(* IEC 61131-3 sources: lasal-git-demo/CPU/LasalDemoProject/Class/ECAT_Master_Base (part 2) *)

#ifdef ECAT_DEBUG_TIMEMEASURE2
          pCTI^.ud_TimePre := OS_GETMICROSEC() - udTimeMarkus;
          if pCTI^.ud_TimePre < pCTI^.ud_TimePreMin then
            pCTI^.ud_TimePreMin := pCTI^.ud_TimePre;
          end_if;
          if pCTI^.ud_TimePre > pCTI^.ud_TimePreMax then
            pCTI^.ud_TimePreMax := pCTI^.ud_TimePre;
          end_if;
#endif
        else

          //Check the process state if we need to raise an error
          dTriggerFrameError := ProcessFrameErrorCheck(pCTI^.ecatm_cycctx^.prcstatus);

          //Check if we need to trigger an error
          if dTriggerFrameError then
            ClassState := _WrongRunStatus;

            bd_LogRtMessagesInCy.PostIt.CycPrcStatus  := TRUE;
            bd_LogRtMessagesInCy.aLogValue1[14]       := pCTI^.ecatm_cycctx^.prcstatus;

            if bd_Flags.bIsRequired then
              CrashThisTime := TRUE;
              sigclib_sprintfST(pd:=#aCrashMessage[0], format:="Ethercat: Error (Invalid frame) Status 0x%X", p0:=#pCTI^.ecatm_cycctx^.prcstatus);
            end_if;
          end_if;
        end_if;

        MissedFrameCounter := sDebugCounters.udConsecutiveMissingFrameCounter;

      end_if;

    else

      sDebugCounters.udInvalidcycctx += 1;

      //Cyclic Context is not valid until EtherCAT State is OP or higher
      if EtherCATState >= ECAT_STATE_OP then
        //Cyclic context is invalid although the EtherCAT State is higher or equal than SAFEOP --> SET Error
        ClassState    := _WrongRunStatus;

        bd_LogRtMessagesInCy.PostIt.InvalidCycctx := TRUE;

        if bd_Flags.bIsRequired then
          CrashThisTime := TRUE;
          _strcpy(dest:=#aCrashMessage[0], src:="EtherCAT: Invalid Cycctx");
        end_if;
      end_if;

    end_if;

  else

    if retcode < ECATM_OK then  // retcode may be of type t_e_st_ecatm_evtc in this case we need unlock
      bNoUnlock := TRUE;
    end_if;

    sDebugCounters.udInvalidRetCodeUpdateCycPre += 1;

    CrashThisTime := UpdateCycRetcodeHandling(retcode:=retcode, pCrashMessage:=#aCrashMessage[0]);

  end_if;

  // Always Call to unlock cycctx
  if ( (pCTI^.bPostScanActive) = FALSE |    // Postscan call needed to unlock ecatm_cycctx
       (EtherCATState < ECAT_STATE_OP) |    // If EtherCATState = OP then unlock is done in postscan
       ((ClassState <> _ClassOk) & (bNoUnlock = FALSE)) ) then     // Unlock on Error, Postscan is no longer called in this state

#ifdef ECAT_TRACE_VIEW_LOG
    OS_MakeTraceEntry(pSystrace, HWCONTROL_SYSTRACE_TYPE, ECAT_SYSTRACE_PRESCAN_UPDATECYC_UNLOCK,pCTI^.udCycTaskId);
#endif

    retcode := OS_ECATM_UpdateCyc(pECAT, ecatmhdl, pCTI^.udCycTaskId, LSL_ECATM_POST_CYC_TASK, #pCTI^.ecatm_cycctx,0);
    if retcode <> ECATM_OK then

      //Invalid retcode, raise error
      sDebugCounters.udInvalidRetCodeUpdateCycPost += 1;

      CrashThisTime := UpdateCycRetcodeHandling(retcode:=retcode, pCrashMessage:=#aCrashMessage[0]);

    end_if;
  end_if;

  if CrashThisTime then
    // if a required module is not available or doesn't work properly, the system should crash
    OS_ECATM_raise_error(pECAT,0,#aCrashMessage[0]);
  end_if;

END_FUNCTION

FUNCTION VIRTUAL GLOBAL ECAT_Master_Base::UpdateRtPostScan
  VAR_INPUT
    pCTI 	: ^t_s_CycTaskInfo;
  END_VAR
  VAR
    i               : UDINT;
    pCallbackData   : ^t_s_MapPDOData;
    CrashThisTime   : BOOL;
    aCrashMessage   : ARRAY [0..255] OF CHAR;
    retcode         : DINT;
    dTriggerFrameError  : DINT;
    prcstatus       : UDINT;
#ifdef ECAT_DEBUG_TIMEMEASURE2
    udTimeMarkus : UDINT;
#endif
  END_VAR

  CrashThisTime   := FALSE; // init with false

  //Check if we have postscan callbacks and a valid frame
  if pCTI^.noPostCallbacks & pCTI^.ecatm_cycctx then

    pCallbackData := pCTI^.pPostCallbacks;
    prcstatus := pCTI^.ecatm_cycctx^.prcstatus; // Save prcstatus as it is checked more than once
    if (prcstatus AND ECATM_PRCSTAT_ST_FRAME_NOT_SENT) = 0 then // ECATM_PRCSTAT_ST_FRAME_NOT_SENT: The link layer driver failed to send the last TX frame.
                                                                //                                  The frame is still owned by the hardware of the MAC.
                                                                //                                  THE APPLICATION SHALL NOT ALTER THE TRANSMIT FRAME!
                                                                // Check the sample-simple and sample-all implementation for usaage and compatibility patch.
                                                                // See ECATM_Programmers_Guide and ECATM_Reference_Manual for detailed information

#ifdef ECAT_DEBUG_TIMEMEASURE2
      udTimeMarkus := OS_GETMICROSEC();
#endif

      //Go through all installed callbacks from the slave modules HWK to fetch the data and copy it to the transmit frame.
      for i := 1 to pCTI^.noPostCallbacks do

        if pCallbackData^.pEtherCatState^ >= ECAT_STATE_OP then

#ifdef ECAT_TRACE_VIEW_LOG
            OS_MakeTraceEntry(pSystrace, HWCONTROL_SYSTRACE_TYPE, ECAT_SYSTRACE_POSTSCAN_CALLBACKS,pCTI^.udCycTaskId OR (i SHL 16));
#endif

          pCallbackData^.pCallBack$ECAT_MapPDOData(pCallbackData^.pThis, pCTI^.ecatm_cycctx, pCallbackData^.noData, pCallbackData^.iovar, pCallbackData^.pData);
        end_if;

        pCallbackData += sizeof(t_s_MapPDOData);
      end_for;

#ifdef ECAT_DEBUG_TIMEMEASURE2
      pCTI^.ud_TimePost := OS_GETMICROSEC() - udTimeMarkus;
      if pCTI^.ud_TimePost < pCTI^.ud_TimePostMin then
        pCTI^.ud_TimePostMin := pCTI^.ud_TimePost;
      end_if;
      if pCTI^.ud_TimePost > pCTI^.ud_TimePostMax then
        pCTI^.ud_TimePostMax := pCTI^.ud_TimePost;
      end_if;
#endif
    end_if;

    if (prcstatus AND ECATM_PRCSTAT_ST_MASK_ERROR_OR_WARN) then

      //Check only if no Prescan is used - otherwise this check is done in prescan
      if pCTI^.noPreCallbacks = 0 then

        //Check the process state if we need to raise an error
        dTriggerFrameError := ProcessFrameErrorCheck(prcstatus);

        if dTriggerFrameError then
          ClassState := _WrongRunStatus;

          bd_LogRtMessagesInCy.PostIt.CycPrcStatus  := TRUE;
          bd_LogRtMessagesInCy.aLogValue1[14]       := prcstatus;

          if bd_Flags.bIsRequired then
            CrashThisTime := TRUE;
            sigclib_sprintfST(pd:=#aCrashMessage[0], format:="Ethercat: Error (Invalid frame) Status 0x%X", p0:=#prcstatus);
          end_if;
        end_if;
      end_if;
    end_if;

    MissedFrameCounter := sDebugCounters.udConsecutiveMissingFrameCounter;

  end_if;

#ifdef ECAT_TRACE_VIEW_LOG
  OS_MakeTraceEntry(pSystrace, HWCONTROL_SYSTRACE_TYPE, ECAT_SYSTRACE_POSTSCAN_UPDATECYC,pCTI^.udCycTaskId);
#endif

  // Always Call to unlock cyctx
  retcode := OS_ECATM_UpdateCyc(pECAT, ecatmhdl, pCTI^.udCycTaskId, LSL_ECATM_POST_CYC_TASK, #pCTI^.ecatm_cycctx,0);

  if udDisconnectEventTime then
    udDisconnectEventTime := 0;
    ClassState := _NoHardware;
    EtherCATState := ECAT_STATE_INIT;
    NewMasterEtherCATState  := ECAT_STATE_INIT;
    InitSSW := _Wait4EcatLink;
  end_if;

  if retcode <> ECATM_OK then
    //Invalid retcode, raise error
    sDebugCounters.udInvalidRetCodeUpdateCycPost += 1;

    CrashThisTime := UpdateCycRetcodeHandling(retcode:=retcode, pCrashMessage:=#aCrashMessage[0]);

  end_if;

  if CrashThisTime then
    // if a required module is not available or doesn't work properly, the system should crash
    OS_ECATM_raise_error(pECAT,0,#aCrashMessage[0]);
  end_if;

END_FUNCTION

FUNCTION VIRTUAL ECAT_Master_Base::UpdateCycRetcodeHandling
  VAR_INPUT
    retcode 	: DINT;
    pCrashMessage : ^Char;
  END_VAR
  VAR_OUTPUT
    bFatalError : BOOL;
  END_VAR

  bFatalError := FALSE;

  //Difference the single errors
  case retcode of
    //*****************************************************************************
    ECATM_TIMING_ERROR_1:

      //No Data available at send time (last cycle)
      ClassState := _TimesliceErrorIRQ;
      bd_LogRtMessagesInCy.PostIt.TimingError_1 := TRUE;

      if bd_Flags.bIsRequired then
        bFatalError := TRUE;
        _strcpy(dest:=pCrashMessage, src:="No Data available at Send time (TimeSliceErrorIRQ)");
      end_if;

    //*****************************************************************************
    ECATM_TIMING_ERROR_2:

      //Time since tick is at call of UpdateCyc(Pre) higher than allowed from the IsoStartPoint
      ClassState := _TimesliceErrorIRQ;
      bd_LogRtMessagesInCy.PostIt.TimingError_2 := TRUE;

      if bd_Flags.bIsRequired then
        bFatalError := TRUE;
        _strcpy(dest:=pCrashMessage, src:="Time since tick is at call of UpdateCyc(Pre) higher than allowed from the IsoStartPoint (TimeSliceErrorIRQ)");
      end_if;

    //*****************************************************************************
    ECATM_DATA_NOT_SENT:

      //Data was not sent at the time UpdateCyc was called with (Pre)
      ClassState := _TimesliceError;
      bd_LogRtMessagesInCy.PostIt.DataNotSent := TRUE;

      if bd_Flags.bIsRequired then
        bFatalError := TRUE;
        _strcpy(dest:=pCrashMessage, src:="Data was not sent at the time UpdateCyc was called with (Pre) (TimeSliceError)");
      end_if;

    //*****************************************************************************
    else

      if retcode = ECATM_EVTC_MST_DEACTIVATED$DINT & InitSSW <> _InitFinished then
        //Ignore master deactivated error during initialisation (maybe master is not activated yet (takes a while in OS)

      else
        ClassState := _ManagerError;
        bd_LogRtMessagesInCy.PostIt.UnknownError := TRUE;
        bd_LogRtMessagesInCy.aLogValue1[4] := (ABS(retcode))$UDINT;
        if bd_Flags.bIsRequired then
          bFatalError := TRUE;
          sigclib_sprintfST(pd:=pCrashMessage, format:="Unknown Error in EtherCAT handling occured: %d", p0:=#retcode);
        end_if;
      end_if;

    //*****************************************************************************
  end_case;

END_FUNCTION

FUNCTION VIRTUAL GLOBAL ECAT_Master_Base::SoftwareVersion::Read
  VAR_OUTPUT
    output (EAX) 	: UDINT;
  END_VAR

  SoftwareVersion := strSoftwareVersion.Data.Read();
  output := SoftwareVersion;

END_FUNCTION

FUNCTION VIRTUAL GLOBAL ECAT_Master_Base::SoftwareVersion::Write
  VAR_INPUT
    input (EAX) 	: UDINT;
  END_VAR
  VAR_OUTPUT
    result (EAX) 	: UDINT;
  END_VAR

  SoftwareVersion := input;
  result := (strSoftwareVersion.Data.Write(SoftwareVersion))$UDINT;

END_FUNCTION

FUNCTION VIRTUAL GLOBAL ECAT_Master_Base::CyWork
  VAR_INPUT
    EAX 	: UDINT;
  END_VAR
  VAR_OUTPUT
    state (EAX) 	: UDINT;
  END_VAR
  VAR
    pCurrentSlave : ^t_sSlaveInfo;
    i             : UDINT;
    _Para         : CmdStruct;
    _Result       : Results;
    RetCodeIPR    : iprStates;
    b_ModulInitComplete   : BOOL;
    TmpRequest    : BDINT;
    retCode       : DINT;
  END_VAR

  case InitSSW of
//**********************************************************************************************************************************************************
    t_e_InitSSW::_StartInit:

#ifdef ECAT_TRACE_VIEW_LOG
      OS_MakeTraceEntry(pSystrace, HWCONTROL_SYSTRACE_TYPE, ECAT_SYSTRACE_POSTINIT_START_INIT,0);
#endif

      // remember when we started (for timeout and init time measure)
      udInitStartTime := ops.tAbsolute;

      // check if we had an error before
      if InitError <> _ClassOk then
        // we already have a log entry from the init
        ClassState := InitError;
        ErrorInitStep := InitSSW;
        InitSSW := _PrepareError;
        EtherCATState := ECAT_STATE_NONE;
        return;
      end_if;

      // Check if post init needs to be extended
      if StateTransitionTimeout.Read() > POST_INIT_TIMEOUT then

        ExtendPostInitTime(AdditionalTime:=StateTransitionTimeout);

      end_if;

      InitSSW := _Wait4ECATLink;

//**********************************************************************************************************************************************************
    t_e_InitSSW::_Wait4ECATLink:

      retCode := OS_ECATM_NET_GET_STATUS(pECAT, ecatmhdl, #snetStatus);

      if retCode then
        LogValue("@0563 (ECAT_Master_Base::CyWork) Failed to get ECAT Link Status. Return Code: 0x{0} via InitModule-Interface", retCode$UDINT);

        ErrorInitStep := InitSSW;
        InitSSW := _PrepareError;
        ClassState := InitError    := _ManagerError;
        EtherCATState := ECAT_STATE_NONE;

        return;
      end_if;

      if snetStatus.flags.ECATM_NET_STATUS_MST_LINK_DOWN = FALSE then

#ifdef ECAT_DEBUG_EVENT_CALLBACKS
        LogValue("ECAT-DEBUG: Link found after 0x{0}ms", (ops.tAbsolute-udInitStartTime));
#endif

        //ClassState is set to NoHardware at DisconnectEvent -> Set back to _ClassOk to ensure that the Realtime functions are called
        ClassState := _ClassOk;

        //Go on and call the connect event methods
        InitSSW := _CallConnectEventOfModules;
      elsif ( (bd_Flags.bDisableWait4LinkTimeOut = FALSE) &
              (ops.tAbsolute - udInitStartTime) > GetWait4LinkTimeout()) then

        ErrorInitStep := InitSSW;
        InitSSW       := _PrepareError;
        ClassState    := InitError     := _ManagerError;
        EtherCATState := ECAT_STATE_NONE;
        LogError("@067B (ECAT_Master_Base::CyWork) Master Link Down (Timeout)! Unable to continue with Initialisation.");

      end_if;

//**********************************************************************************************************************************************************
    t_e_InitSSW::_CallConnectEventOfModules:

      //Call the Connect Event of every slave
      if sSlaveInfo.udMaxSlaves then
        pCurrentSlave := sSlaveInfo.pSlaves; //Point to current slave
        for i:=0 to sSlaveInfo.udMaxSlaves-1 do
          //Only call module if no error
          if pCurrentSlave^.pThis & pCurrentSlave^.pThis^.EtherCATState <> ECAT_STATE_NONE then
            pCurrentSlave^.pThis^.ConnectEvent();
          end_if;
          pCurrentSlave += sizeof(t_sSlaveInfo);
        end_for;
      end_if;

      InitSSW := _PrepareNextEtherCATState;

//**********************************************************************************************************************************************************
    t_e_InitSSW::_PrepareNextEtherCATState:

      //Go on with next step of initialisation
      InitSSW := _SwitchToNextEtherCATState;
      TmpRequest := 0;

      //Check if any slave needs an InitModule call. Otherwise we can directy request the OP State from the master
      if sSlaveInfo.udMaxSlaves then
        pCurrentSlave := sSlaveInfo.pSlaves; //Point to current slave
        //Call UpdateCy of all logged in slaves
        for i:=0 to sSlaveInfo.udMaxSlaves-1 do
          if pCurrentSlave^.pThis & pCurrentSlave^.bdInitModuleFlags <> ECAT_INIT_MODULE_NO_CALL then
            TmpRequest := TmpRequest OR pCurrentSlave^.bdInitModuleFlags;
          end_if;
          pCurrentSlave += sizeof(t_sSlaveInfo);
        end_for;
      end_if;

      //Determine master state to request (e.g. if no module needs to be called during our InitModulePhase, we can directly request the OP State)
      if (TmpRequest AND ECAT_INIT_MODULE_CALL_INIT) = ECAT_INIT_MODULE_CALL_INIT then
        RequestMasterState := ECAT_STATE_INIT;
      elsif (TmpRequest AND ECAT_INIT_MODULE_CALL_PREOP) = ECAT_INIT_MODULE_CALL_PREOP then
        RequestMasterState := ECAT_STATE_PREOP;
      elsif (TmpRequest AND ECAT_INIT_MODULE_CALL_SAFEOP) = ECAT_INIT_MODULE_CALL_SAFEOP then
        RequestMasterState := ECAT_STATE_SAFEOP;
      else
        //No module needs an InitModule Call
        RequestMasterState := ECAT_STATE_OP;
      end_if;

//**********************************************************************************************************************************************************
    t_e_InitSSW::_SwitchToNextEtherCATState:

      //Set master to determined state
#ifdef ECAT_DEBUG_EVENT_CALLBACKS
      LogValue(pString:="ECAT-DEBUG: Request New ECATMST State: 0x{0}", Value:=RequestMasterState);
#endif
      retcode := OS_ECATM_MST_REQ_STATE(pECAT, ecatmhdl, RequestMasterState, StateTransitionBehaviour);
      if retcode then
        LogValue("@0565 (ECAT_Master_Base::CyWork) Call OS_ECATM_MST_REQ_STATE() Failed with retcode 0x{0}! Unable to continue with Initialisation", ABS(retcode)$UDINT);
        // Disable Class
        ErrorInitStep := InitSSW;
        InitSSW := _PrepareError;
        ClassState := _ManagerError;
        EtherCATState := ECAT_STATE_NONE;
        return;
      end_if;

      udCheckEtherCATStateTime := ops.tAbsolute;
      InitSSW := _CheckEtherCATState;

//**********************************************************************************************************************************************************
    t_e_InitSSW::_CheckEtherCATState:

      //Wait until master is in requested state
      if EtherCATState = RequestMasterState then

#ifdef ECAT_TRACE_VIEW_LOG
        OS_MakeTraceEntry(pSystrace, HWCONTROL_SYSTRACE_TYPE, ECAT_SYSTRACE_POSTINIT_CHECK_ETHERCAT_STATE,EtherCATState$UDINT);
#endif

        //If we are in the requested state go on with InitModule Phase
        InitSSW := _CallInitModule;

        udInitModuleTimeStamp := ops.tAbsolute;
        udInitModuleTimeOut   := GetCallInitModuleTimeout();

      elsif ( (bd_Flags.bDisableStateTransitionTimeout = FALSE) &
              (ops.tAbsolute - udCheckEtherCATStateTime) > StateTransitionTimeout.Read()) then
        LogValue("@0566 (ECAT_Master_Base::CyWork) Timeout while waiting for EtherCATState! EtherCATState: 0x{0}, RequestMasterState: 0x{1}", EtherCATState$UDINT,RequestMasterState$UDINT);
        ErrorInitStep := InitSSW;
        InitSSW := _PrepareError;
        ClassState := _TimeoutInInit;
        EtherCATState := ECAT_STATE_NONE;
        return;
      end_if;

//**********************************************************************************************************************************************************
    t_e_InitSSW::_CallInitModule:

      // preinitialize the complete marker => is resetted if a module has to be initialized
      b_ModulInitComplete := TRUE;

      //Call all slaves (needed for SDO Handling)
      if sSlaveInfo.udMaxSlaves then
        pCurrentSlave := sSlaveInfo.pSlaves; //Point to current slave

        _Para.uiCmd := ECAT_M_CALL_INIT_MODULE;
        _Para.aPara[0]$DINT           := 1;
        _Para.aPara[1]$t_e_ECAT_STATE := EtherCATState;

        //Call UpdateCy of all logged in slaves
        for i:=0 to sSlaveInfo.udMaxSlaves-1 do

          //Check if current module has to be called
          if (pCurrentSlave^.bdInitModuleFlags <> ECAT_INIT_MODULE_NO_CALL) &
            ((pCurrentSlave^.bdInitModuleFinished AND EtherCATState$BDINT) <> EtherCATState$BDINT ) then

            if (EtherCATState = ECAT_STATE_INIT   & ((pCurrentSlave^.bdInitModuleFlags AND ECAT_INIT_MODULE_CALL_INIT)    = ECAT_INIT_MODULE_CALL_INIT))  |
               (EtherCATState = ECAT_STATE_PREOP  & ((pCurrentSlave^.bdInitModuleFlags AND ECAT_INIT_MODULE_CALL_PREOP)   = ECAT_INIT_MODULE_CALL_PREOP)) |
               (EtherCATState = ECAT_STATE_SAFEOP & ((pCurrentSlave^.bdInitModuleFlags AND ECAT_INIT_MODULE_CALL_SAFEOP)  = ECAT_INIT_MODULE_CALL_SAFEOP)) |
               (EtherCATState = ECAT_STATE_OP     & ((pCurrentSlave^.bdInitModuleFlags AND ECAT_INIT_MODULE_CALL_OP)      = ECAT_INIT_MODULE_CALL_OP))
            then
              RetCodeIPR := pCurrentSlave^.pThis^.NewInst(#_Para,#_Result);

#ifdef ECAT_TRACE_VIEW_LOG
              OS_MakeTraceEntry(pSystrace, HWCONTROL_SYSTRACE_TYPE, ECAT_SYSTRACE_POSTINIT_CALL_INITMODULE,i);
#endif
              //Check retcode
              if RetCodeIPR = ERROR then

                LogValue("@0567 (ECAT_Master_Base::CyWork) Failed to initialize EtherCAT Slave 0x{0} via InitModule-Interface", i);

                // Set as finshed so that not required module is not called again and does not spam log
                // Disable Init callbacks for all EtherCAT States
                pCurrentSlave^.bdInitModuleFinished := pCurrentSlave^.bdInitModuleFinished OR ECAT_STATE_INIT$BDINT OR ECAT_STATE_PREOP$BDINT OR ECAT_STATE_SAFEOP$BDINT OR ECAT_STATE_OP$BDINT;

                // if it's an required module => error
                if pCurrentSlave^.bRequired   then
                  SetRequiredError( pTargetThis       := pCurrentSlave^.pThis
                                  , udSlaveIndex      := pCurrentSlave^.udSlaveIndex
                                  , bLogInMethAllowed := TRUE);
                end_if;

              elsif RetCodeIPR = READY then
                pCurrentSlave^.bdInitModuleFinished := pCurrentSlave^.bdInitModuleFinished OR EtherCATState$BDINT;
              else
                b_ModulInitComplete := FALSE; //At least one module is not ready yet --> carry on with ModuleInit phase
              end_if;
            //else
              //Module will be called if the needed EtherCAT State is active
            end_if;
          else
            //Module has no need to be called, just set as finished
            pCurrentSlave^.bdInitModuleFinished := pCurrentSlave^.bdInitModuleFinished OR EtherCATState$BDINT;
          end_if;

          pCurrentSlave += sizeof(t_sSlaveInfo);
        end_for;
      end_if;

      //Check if every module init is finished, go on to next state
      if b_ModulInitComplete = TRUE then

        InitSSW := _SwitchToNextEtherCATState;

        case EtherCATState of
        //*****************************************************************************
          t_e_ECAT_STATE::ECAT_STATE_INIT:
            //Next step to request is Preop
            RequestMasterState := ECAT_STATE_PREOP;

        //*****************************************************************************
          t_e_ECAT_STATE::ECAT_STATE_PREOP:
            //Next step to request is SafeOP
            RequestMasterState := ECAT_STATE_SAFEOP;

        //*****************************************************************************
          t_e_ECAT_STATE::ECAT_STATE_SAFEOP:

            // Configure Synchronisation ***********************************************************************
            if ( (sDCInfo.DCModuleEnabled) &                  // Only when DC unit is enabled
                 (sDCInfo.SyncMeasureConfigOk = FALSE) ) then
              if Config_SyncMeasureECAT() <> ECAT_RETOK then
                SetRequiredError(bLogInMethAllowed := TRUE);
              end_if;
            end_if;
            // Configure Synchronisation end ********************************************************************

            //Next step to request is OP
            RequestMasterState := ECAT_STATE_OP;

        //*****************************************************************************
          t_e_ECAT_STATE::ECAT_STATE_OP:

            //Finished, check if we have a DC Module --> we need to wait until everything is synchron
            if sDCInfo.DCModuleEnabled = TRUE then

              // Configure Synchronisation ***********************************************************************
              // Check again incase SAFE_OP was skipped
              if (sDCInfo.SyncMeasureConfigOk = FALSE) then
                if Config_SyncMeasureECAT() <> ECAT_RETOK then
                  SetRequiredError(bLogInMethAllowed := TRUE);
                end_if;
              end_if;
              // Configure Synchronisation end ********************************************************************
              InitSSW := _WaitForSynchron;
              udWaitForSynchronTimeStamp := ops.tAbsolute;
            else
              InitSSW := _FinishInitialisation;
            end_if;

            udTimeUntilOP := ops.tAbsolute - udInitStartTime;

        //*****************************************************************************

        end_case;

      elsif (bd_Flags.bDisableInitModuleTimeOut = FALSE) &
            (ops.tAbsolute - udInitModuleTimeStamp) > udInitModuleTimeOut then
        LogError("@0568 (ECAT_Master_Base::CyWork) Timeout in CallInitModule step.");
        ErrorInitStep := InitSSW;
        InitSSW := _PrepareError;
        ClassState := _TimeoutInInit;
        EtherCATState := ECAT_STATE_NONE;
        return;
      end_if;

//**********************************************************************************************************************************************************
    t_e_InitSSW::_WaitForSynchron: //Wait until synchron

      //Wait until class is synchron
      if _SyncMeasureECAT1.Synchron then
#ifdef ECAT_TRACE_VIEW_LOG
        OS_MakeTraceEntry(pSystrace, HWCONTROL_SYSTRACE_TYPE, ECAT_SYSTRACE_POSTINIT_IS_SYNCRHON,0);
#endif
        udTimeSynchron := ops.tAbsolute - udTimeUntilOP + udInitStartTime;
        InitSSW := _FinishInitialisation;

      elsif ( (bd_Flags.bDisableWaitForSynchronTimeOut = FALSE) &
              ((ops.tAbsolute - udWaitForSynchronTimeStamp) > GetWait4SynchronTimeout()) ) then
        LogError("@0569 (ECAT_Master_Base::CyWork) Timeout while waiting for synchron");
        ErrorInitStep := InitSSW;
        InitSSW := _PrepareError;
        ClassState := _TimeoutInInit;
        EtherCATState := ECAT_STATE_NONE;
        return;
      end_if;

//**********************************************************************************************************************************************************
    t_e_InitSSW::_FinishInitialisation:

      //we're finished with initializing
      bd_Flags.bPostInitFinished := TRUE;

      udInitDuration := ops.tAbsolute - udInitStartTime;

#ifdef ECAT_TRACE_VIEW_LOG
      OS_MakeTraceEntry(pSystrace, HWCONTROL_SYSTRACE_TYPE, ECAT_SYSTRACE_POSTINIT_INIT_FINISHED,0);
#endif

      InitSSW := _InitFinished;

//**********************************************************************************************************************************************************
    t_e_InitSSW::_InitFinished: //Normal cyclic work

      if ClassState <> _ClassOk then

        // Error occoured at EtherCat Master
        // Sets Slaves into error state
        SendManagerErrorToSlaves();

        InitSSW := _PrepareError;

      end_if;

//**********************************************************************************************************************************************************
    t_e_InitSSW::_PrepareError: // do error handling and then stay in _ErrorOccured-Step

      //we're finished with initializing
      bd_Flags.bPostInitFinished := TRUE;
      InitSSW := _ErrorOccured;

      if bd_Flags.bIsRequired then
        SetRequiredError(bLogInMethAllowed := TRUE);
      else
        // The following code switches off the BUS completely.
        // Advantage: No subsequent errors because HWK is deactivated. Disadvantage: SDOs for diagnostics are disabled!
        // For the SDOs part of the Rt must continue to run, otherwise the EtherCAT states will no longer function correctly. see OS_ECATM_UpdateCyc
        DisconnectEvent(udMasterID:=0, evt:=NIL, EventType:=0, uiCallbackInfo:=0);
        // Deactivate Master
        StartChangeMasterState(FALSE);
        InitSSW := _ErrorOccuredWait4MasterDeactivate;
      end_if;

//**********************************************************************************************************************************************************
    t_e_InitSSW::_ErrorOccuredWait4MasterDeactivate:

      if GetStateChangeMasterState() <> BUSY then
        InitSSW := _ErrorOccured;
      end_if;

//**********************************************************************************************************************************************************
    t_e_InitSSW::_ErrorOccured: // do nothing here
      //return; //No return here otherwise realtime log messages will not be logged anymore

//**********************************************************************************************************************************************************
    t_e_InitSSW::_NotConnected:

      // Disable Syncregulation if active
      if _SyncMeasureECAT1.SyncRegulationEnable then
        _SyncMeasureECAT1.SyncRegulationEnable.Write(input:=0);
        sDCInfo.SyncMeasureConfigOk := FALSE;
      end_if;

  end_case;

  //Always call all slaves (needed for SDO Handling)
  if sSlaveInfo.udMaxSlaves then
    pCurrentSlave := sSlaveInfo.pSlaves; //Point to current slave
    //Call UpdateCy of all logged in slaves
    for i:=0 to sSlaveInfo.udMaxSlaves-1 do

      //Check if slave should be called
      if pCurrentSlave^.pThis & pCurrentSlave^.pThis^.EtherCATState <> ECAT_STATE_NONE then
        pCurrentSlave^.pThis^.UpdateCy();
      end_if;

      pCurrentSlave += sizeof(t_sSlaveInfo);
    end_for;
  end_if;

  // Call for loggin
  _SyncMeasureECAT1.CyWork(EAX:=0);

  //Log messages from realtime in cyclic
  LogRtMessages();

  state := READY;

END_FUNCTION

FUNCTION ECAT_Master_Base::StartChangeMasterState
	VAR_INPUT
		EnableMasterState 	: BOOL;
	END_VAR
	VAR_OUTPUT
		retcode 	: iprStates;
	END_VAR
  VAR
	  astr_threadname : ARRAY [0..30] OF CHAR;
  END_VAR

  retcode := BUSY;

  if (sChangeMasterState.bdFlags.TaskActivated = FALSE) & (sChangeMasterState.bdFlags.TaskActive = FALSE) then  // Only start thread if not active

    sChangeMasterState.bdFlags.TaskDone      := FALSE;
    sChangeMasterState.bdFlags.TaskActivated := TRUE;

    sChangeMasterState.bdFlags.EnableMaster := EnableMasterState;

    //Create a dynamic threadname
    sigclib_strcpy(#astr_threadname[0], "ChangeMasterStateHndl");
    sigclib_htoa(#astr_threadname[sigclib_strlen(#astr_threadname[0])], this$udint);

    // Needs own thread because OS call is blocking
    sChangeMasterState.mtTaskHandle := toMultiTask.CREATETHREAD(taskfunction0 := #ChangeMasterState()
                                                              , priority0     := ECATM_THREAD_PRIO_DISABLE   // priority same as background
                                                              , stackSize0    := ECATM_THREAD_STACKSIZE
                                                              , flags0        := MT_TASK_SAVETHIS
                                                              , parameter0    := THIS
                                                              , name0         := #astr_threadname[0]);

    retcode := READY;

  end_if;

END_FUNCTION

FUNCTION ECAT_Master_Base::GetStateChangeMasterState
	VAR_OUTPUT
		retcode 	: iprStates;
	END_VAR

  retcode := BUSY;
  if (sChangeMasterState.bdFlags.TaskActivated = FALSE) & (sChangeMasterState.bdFlags.TaskActive = FALSE) then
    retcode := READY;
  end_if;

END_FUNCTION

FUNCTION ECAT_Master_Base::ChangeMasterState

  sChangeMasterState.bdFlags.TaskActive    := TRUE;
  sChangeMasterState.bdFlags.TaskActivated := FALSE;

  sChangeMasterState.retcode := OS_ECATM_MASTER_ACTIVATE(pECAT, ecatmhdl, sChangeMasterState.bdFlags.EnableMaster);

  sChangeMasterState.bdFlags.TaskDone   := TRUE;
  sChangeMasterState.bdFlags.TaskActive := FALSE;

END_FUNCTION

FUNCTION VIRTUAL GLOBAL ECAT_Master_Base::Synchron::Read
  VAR_OUTPUT
    output (EAX) 	: DINT;
  END_VAR

  Synchron := _SyncMeasureECAT1.Synchron.Read();
  output := Synchron;

END_FUNCTION

FUNCTION VIRTUAL ECAT_Master_Base::Config_SyncMeasureECAT
	VAR_OUTPUT
		retcode 	: DINT;
	END_VAR
  VAR
    _Para 	      : CmdStruct;
    _Result 	    : Results;
    ret_code 	    : IprStates;
    pCurrentSlave : ^t_sSlaveInfo;
    i             : UDINT;
    pCTI          : ^t_s_CycTaskInfo;
    bcycidxOk     : BOOL;
  END_VAR

  // Get ECAT Bus period (must be called in state SAFEOP or higher)
  retcode := OS_ECATM_DC_GET_STATS(pECAT, ecatmhdl, #sDC_Stats);

  if retcode then
    LogValue("@056A (ECAT_Master_Base::Config_SyncMeasureECAT) Call OS_ECATM_dc_get_stats() Failed with retcode: {0}!", retcode$UDINT);
  else

    retcode := ECAT_RETERR_CMD_INVALID_SLV;
    if sSlaveInfo.udMaxSlaves >= sDCInfo.udSlaveIndex then
      pCurrentSlave := sSlaveInfo.pSlaves + (sDCInfo.udSlaveIndex * sizeof(t_sSlaveInfo) );

      if pCurrentSlave^.pThis then

        // Get Cycidx from DC Slave
        _Para.uiCmd     := ECAT_M_GET_SLAVE_CYCIDX;
        _Para.aPara[0]  := 1; // Version

        ret_code := pCurrentSlave^.pThis^.NewInst(#_Para,#_Result);
        retcode := ECAT_RETERR_CMD_CYCIDX_NOTFOUND;
        if (ret_code = READY) & (_Result.uiLng = 12) &
           (_Result.aData[0]$DINT = ECAT_RETOK) &
           (_Result.aData[4]$DINT = 1) then // Version

          sDCInfo.udCyclicIndex :=  _Result.aData[8];

          // Search Cycle task for the tasks in which the DC time is received
          i         := 0;
          bcycidxOk := FALSE;
          pCTI      := pCycTaskInfo;
          while i < udNoCycTasks do

            if pCTI^.udCycTaskId = sDCInfo.udCyclicIndex then

              // _SyncMeasureECAT1.Set_PeriodTimeMaster((sDC_Stats.cyctime * 1000)$DINT ); // *1000 us => ns

              _SyncMeasureECAT1.Set_PeriodTimeMaster((pCTI^.udCycleTime_us * 1000)$DINT ); // *1000 us => ns

              // Start synchrone data
              _SyncMeasureECAT1.Set_PeriodTimeOwn(newPeriodTimeOwn := (pCTI^.udCycleTime_us * 1000)$DINT );

              if bs_syncmodes.DCSlavemodeActive then
                _SyncMeasureECAT1.SyncRegulationEnable.Write(input:=1);//The ECAT DC will be adjusted
              else
                _SyncMeasureECAT1.SyncRegulationEnable.Write(input:=2);//The Sigmatek PLL will be adjusted
              end_if;

              bcycidxOk := TRUE;
              sDCInfo.SyncMeasureConfigOk := TRUE;
              retcode := ECAT_RETOK;
              exit;
            end_if;

            i += 1;
            pCTI += sizeof(t_s_CycTaskInfo);

          end_while;

          if bcycidxOk = FALSE then
            LogValue("@056B (ECAT_Master_Base::Config_SyncMeasureECAT) Failed to find sDCInfo.cycidx: 0x{0}!", sDCInfo.udCyclicIndex);
          end_if;
        else
          LogValue("@056C (ECAT_Master_Base::Config_SyncMeasureECAT) NewInstCmd: ECAT_M_GET_SLAVE_CYCIDX Failed! ret_code = 0x{0}, return code = 0x{1}, Version = 0x{2}", ret_code$UDINT, _Result.aData[0]$UDINT, _Result.aData[4]$UDINT);
        end_if;

      else  // if pCurrentSlave^.pThis then
        LogValue("@056D (ECAT_Master_Base::Config_SyncMeasureECAT) Invalid sDCInfo.slvidx: 0x{0}!", sDCInfo.udSlaveIndex);
      end_if;

    else  // if sSlaveInfo.udMaxSlaves >= sDCInfo.udSlaveIndex then
      LogValue("@056F (ECAT_Master_Base::Config_SyncMeasureECAT) Invalid sDCInfo.slvidx: 0x{0}!", sDCInfo.udSlaveIndex);
    end_if;
  end_if;

END_FUNCTION

FUNCTION VIRTUAL ECAT_Master_Base::LogRtMessages
  VAR
  	bPostIt : t_b_RtMessages;
  END_VAR

  // if there are some messages to post, post them (the methods in the brackets are not the actual, but the methods were the error occured)
  if bd_LogRtMessagesInCy.PostIt then

    bPostIt := bd_LogRtMessagesInCy.PostIt;

    if bPostIt.InvalidNewInstCommandReceived  then
      LogValue("@0570 (ECAT_Master_Base::EtherCATState::NewInst) Received unknown command: 0x{0}", bd_LogRtMessagesInCy.aLogValue1[0]);
    end_if;

    if bPostIt.UnknownCallbackReceived  then
      LogValue("@0571 (ECAT_Master_Base::EtherCATState::NewInst) Received unknown callback: 0x{0}", bd_LogRtMessagesInCy.aLogValue1[1]);
    end_if;

    if bPostIt.UnknownError  then
      LogValue("@0574 (ECAT_Master_Base::UpdateRt) Unknown Error occured: 0x{0}", bd_LogRtMessagesInCy.aLogValue1[4]);
    end_if;

    if bPostIt.SlvTransFailed then
      LogValue("@0575 (ECAT_Master_Base::EvtCallBack) State transition of required Slave 0x{0} failed.", bd_LogRtMessagesInCy.aLogValue1[5]);
    end_if;

    if bPostIt.SendEvtCallInvSlv then
      LogValue("@0576 (ECAT_Master_Base::SendEvtCallBacktoSlave) Invalid slave number from Event callback! evt^.arg1 = 0x{0}", bd_LogRtMessagesInCy.aLogValue1[6]);
    end_if;

    if bPostIt.SendEvtCallInvFailed then
      LogValue("@0577 (ECAT_Master_Base::SendEvtCallBacktoSlave) NewInstCmd: ECAT_M_EVENT_CALLBACK Failed! return code = 0x{0}, Version = 0x{2}", bd_LogRtMessagesInCy.aLogValue1[7]);
    end_if;

    if bPostIt.SetReqErrSlv then
      LogValue("@0579 (ECAT_Master_Base::SetRequiredError) Required Error on EtherCAT Slave 0x{0}.", bd_LogRtMessagesInCy.aLogValue1[8] );
    end_if;

    if bPostIt.SetReqErrFailed then
      LogError("@057A (ECAT_Master_Base::SetRequiredError) Failed to raise Required Error.");
    end_if;

    if bPostIt.InitCRecvTimeout then
      LogValue("@057B (ECAT_Master_Base::EvtCallBack) Init command failed with frame timeout error. Device Index: 0x{0}",bd_LogRtMessagesInCy.aLogValue1[10]);
    end_if;

    if bPostIt.InitCValidWKC then
      LogValue("@057C (ECAT_Master_Base::EvtCallBack) Init command failed failed with wrong working counter. Device Index: 0x{0}",bd_LogRtMessagesInCy.aLogValue1[11]);
    end_if;

    if bPostIt.InitCValidLen then
      LogValue("@09C8 (ECAT_Master_Base::EvtCallBack) Init command failed with invalid frame length. Device Index: 0x{0}",bd_LogRtMessagesInCy.aLogValue1[12]);
    end_if;

    if bPostIt.InitCValidData then
      LogValue("@057E (ECAT_Master_Base::EvtCallBack) Init command failed during data validation. Device Index: 0x{0}",bd_LogRtMessagesInCy.aLogValue1[13]);
    end_if;

    if bPostIt.CycPrcStatus & bd_LogRtMessagesInCy.AlreadyPosted.CycPrcStatus = FALSE then
      LogValue("@057F (ECAT_Master_Base::UpdateRt) Invalid status of cyclic context detected: prcstatus: 0x{0}",bd_LogRtMessagesInCy.aLogValue1[14]);
      bd_LogRtMessagesInCy.AlreadyPosted.CycPrcStatus := TRUE;
    end_if;

    if bPostIt.DCSlaveTransFailed then
      LogValue("@0580 (ECAT_Master_Base::EvtCallBack) State transition of DC Slave 0x{0} failed.", bd_LogRtMessagesInCy.aLogValue1[15]);
    end_if;

    if bPostIt.InvalidDCCyclePeriod then
      LogValue("@0581 (ECAT_Master_Base::EvtCallBack) Sync0 period of the slave 0x{0} is not a multiple or fraction of the cyclic task period",bd_LogRtMessagesInCy.aLogValue1[16]);
    end_if;

    if bPostIt.NoFreeReceiveFrameBuffer & bd_LogRtMessagesInCy.AlreadyPosted.NoFreeReceiveFrameBuffer = FALSE then
      LogError("@0583 (ECAT_Master_Base::EvtCallBack) No free receive frame buffer (check ecatm configuration)");
      bd_LogRtMessagesInCy.AlreadyPosted.NoFreeReceiveFrameBuffer := TRUE;
    end_if;

    if bPostIt.InvalidCycctx & bd_LogRtMessagesInCy.AlreadyPosted.InvalidCycctx = FALSE then
      LogError("@0922 (ECAT_Master_Base::UpdateRt) Invalid Cycctx");
      bd_LogRtMessagesInCy.AlreadyPosted.InvalidCycctx := TRUE;
    end_if;

    if bPostIt.TimingError_1 & bd_LogRtMessagesInCy.AlreadyPosted.TimingError_1 = FALSE then
      LogError("@0923 (ECAT_Master_Base::UpdateRt) No Data available at Send time (TimeSliceErrorIRQ)");
      bd_LogRtMessagesInCy.AlreadyPosted.TimingError_1 := TRUE;
    end_if;

    if bPostIt.TimingError_2 & bd_LogRtMessagesInCy.AlreadyPosted.TimingError_2 = FALSE then
      LogError("@0924 (ECAT_Master_Base::UpdateRt) Time since tick is at call of UpdateCyc(Pre) higher than allowed from the IsoStartPoint (TimeSliceErrorIRQ)");
      bd_LogRtMessagesInCy.AlreadyPosted.TimingError_2 := TRUE;
    end_if;

    if bPostIt.DataNotSent & bd_LogRtMessagesInCy.AlreadyPosted.DataNotSent = FALSE then
      LogError("@0925 (ECAT_Master_Base::UpdateRt) Data was not sent at the time UpdateCyc was called with (Pre) (TimeSliceError)");
      bd_LogRtMessagesInCy.AlreadyPosted.DataNotSent := TRUE;
    end_if;

    bd_LogRtMessagesInCy.PostIt := bd_LogRtMessagesInCy.PostIt AND (NOT bPostIt); // Only delete flags of messages that were posted this time.
  end_if;

#ifdef ECAT_DEBUG_FRAMETIME
  if gavg_FrameTime >= gErrorLimitFT then
    ((0)$^USINT)^ := 0;
    OS_ReportTraceEvent(pSystrace, TEVENT_USER0);
  end_if;
#endif

END_FUNCTION

FUNCTION __CDECL VIRTUAL ECAT_Master_Base::EvtCallBack
	VAR_INPUT
		udMasterID 	: UDINT;
		evt 	: ^t_st_ecatm_evt;
		EventType 	: DINT;
		uiCallbackInfo 	: UINT;
	END_VAR
  VAR
    pCurrentSlave : ^t_sSlaveInfo;
    bLogInCallbackAllowed : BOOL;   //Shows if logging is allowed in the callback
  END_VAR

  //Default: Log in callback is not allowed
  bLogInCallbackAllowed := FALSE;
  //Check if we are getting called from the acyclic task --> we are allowed to log in the callback (no log if we are called in realtime to avoid RtRuntime Error)
  if (uiCallbackInfo = LSL_ECATM_ACYCLIC_TASK) then
    bLogInCallbackAllowed := TRUE;
  end_if;

  //Check for valid event code
  if ( (evt^.evtcode > ECATM_EVTC_FIRST) & (evt^.evtcode < ECATM_EVTC_LAST) ) then
    aCntCallBacks[evt^.evtcode] += 1;
    aCntCallBacks[ECATM_EVTC_LAST] += 1; // Use Last index for global cnt
  else
    //We received an unknown event
    udUnknownEventCallback += 1;

    if bLogInCallbackAllowed = FALSE THEN
      //Log in cyclic
      bd_LogRtMessagesInCy.aLogValue1[1] := (evt^.evtcode)$UDINT;
      bd_LogRtMessagesInCy.PostIt.UnknownCallbackReceived := TRUE;
    else
      HWC_LogPrintf(pThis:=this, format:="@0571 (ECAT_Master_Base::EvtCallBack) Received unknown callback: %V4", #evt^.evtcode);
      HWC_LogPrintf(pThis:=this, format:="@0571 arg1: %d, arg2: %d, arg3: %d, arg4: %d", #evt^.arg1, #evt^.arg2, #evt^.arg3, #evt^.arg4);
    end_if;
  end_if;

#ifdef ECAT_TRACE_VIEW_LOG
  OS_MakeTraceEntry(pSystrace, HWCONTROL_SYSTRACE_TYPE, ECAT_SYSTRACE_POSTINIT_EVTCALLBACK,evt^.evtcode$UDINT);
#endif

  case evt^.evtcode of
//*******************************************************************************************************************************************************
    ECATM_EVTC_BUSY:
    //Function can currently not be performed. Try again.

#ifdef ECAT_DEBUG_EVENT_CALLBACKS
      LogError("ECAT-DEBUG: Function can currently not be performed. Try again");
#endif

//*******************************************************************************************************************************************************
    ECATM_EVTC_ERR_PARAM:
    //Wrong parameter value

#ifdef ECAT_DEBUG_EVENT_CALLBACKS
      LogError("ECAT-DEBUG: Wrong parameter value");
#endif

//*******************************************************************************************************************************************************
    ECATM_EVTC_ERR_BUFSIZE:
    //Buffer size is too small

#ifdef ECAT_DEBUG_EVENT_CALLBACKS
      LogError("ECAT-DEBUG: Buffer size is too small");
#endif

//*******************************************************************************************************************************************************
    ECATM_EVTC_ERR_NOT_SUPPORTED:
    //Operation is not supported

#ifdef ECAT_DEBUG_EVENT_CALLBACKS
      LogError("ECAT-DEBUG: Operation is not supported");
#endif

//*******************************************************************************************************************************************************
    ECATM_EVTC_ERR_TIMEOUT:
    //Timeout error

#ifdef ECAT_DEBUG_EVENT_CALLBACKS
      LogError("ECAT-DEBUG: Timeout error");
#endif

//*******************************************************************************************************************************************************
    ECATM_EVTC_MEM_ALLOC:
    //Memory allocation failed

#ifdef ECAT_DEBUG_EVENT_CALLBACKS
      LogError("ECAT-DEBUG: Memory allocation failed");
#endif

//*******************************************************************************************************************************************************
    ECATM_EVTC_ENI_ERR:
    //Error during ENI parsing (see eceni_file.h)

#ifdef ECAT_DEBUG_EVENT_CALLBACKS
      LogError("ECAT-DEBUG: Error during ENI parsing (see eceni_file.h) ");
#endif

//*******************************************************************************************************************************************************
    ECATM_EVTC_ENI_WARN:
    //Warning during ENI parsing (see eceni_file.h)

#ifdef ECAT_DEBUG_EVENT_CALLBACKS
      LogError("ECAT-DEBUG: Warning during ENI parsing (see eceni_file.h) ");
#endif

//*******************************************************************************************************************************************************
    ECATM_EVTC_CYC_PRCSTATUS_CHG:
    //Cyclic process status changed

#ifdef ECAT_DEBUG_EVENT_CALLBACKS
      LogValue(pString:="ECAT-DEBUG: Cyclic process status changed. New status 0x{0}, Old status 0x{1} ", Value:= evt^.arg2$t_stb_ecatm_prcstat, Value2 := lastPRCStatus);
#endif

    if ( (lastPRCStatus.LINK_ERROR = TRUE) &
         (evt^.arg2$t_stb_ecatm_prcstat.LINK_ERROR = FALSE) ) then
#ifdef ECAT_DEBUG_EVENT_CALLBACKS
      LogError("ECAT-DEBUG: New Link found.");
#endif
      ConnectEvent(udMasterID, evt, EventType, uiCallbackInfo);

    end_if;

    lastPRCStatus := evt^.arg2$t_stb_ecatm_prcstat;

//*******************************************************************************************************************************************************
    ECATM_EVTC_CYC_NOT_DESTROYED:
    //At least one cyclic task is not destroyed

#ifdef ECAT_DEBUG_EVENT_CALLBACKS
      LogError("ECAT-DEBUG: At least one cyclic task is not destroyed");
#endif

//*******************************************************************************************************************************************************
    ECATM_EVTC_CYC_ERR_NO_RCV_TS:
    //The receive time stamp was not provided by the link layer or is marked as invalid.

#ifdef ECAT_DEBUG_EVENT_CALLBACKS
      LogError("ECAT-DEBUG: The receive time stamp was not provided by the link layer or is marked as invalid.");
#endif

//*******************************************************************************************************************************************************
    ECATM_EVTC_CYC_ERR_NO_SND_TS:
    //The send time stamp was not provided by the link layer or is marked as invalid.

#ifdef ECAT_DEBUG_EVENT_CALLBACKS
      LogError("ECAT-DEBUG: The send time stamp was not provided by the link layer or is marked as invalid.");
#endif

//*******************************************************************************************************************************************************
    ECATM_EVTC_IOVAR_BAD_CFG:
    //Process variable configuration does not match to the function

#ifdef ECAT_DEBUG_EVENT_CALLBACKS
      LogError("ECAT-DEBUG: Process variable configuration does not match to the function ");
#endif

//*******************************************************************************************************************************************************
    ECATM_EVTC_IOVAR_BAD_ID:
    //iovarid is invalid

#ifdef ECAT_DEBUG_EVENT_CALLBACKS
      LogError("ECAT-DEBUG: iovarid is invalid");
#endif

//*******************************************************************************************************************************************************
    ECATM_EVTC_IOVAR_BAD_PDO:
    //iovarpdo is invalid

#ifdef ECAT_DEBUG_EVENT_CALLBACKS
      LogError("ECAT-DEBUG: iovarpdo is invalid");
#endif

//*******************************************************************************************************************************************************
    ECATM_EVTC_IOVAR_BAD_NAME:
    //iovarname is invalid

#ifdef ECAT_DEBUG_EVENT_CALLBACKS
      LogError("ECAT-DEBUG: iovarname is invalid");
#endif

//*******************************************************************************************************************************************************
    ECATM_EVTC_IOVAR_BAD_CYCIDX:
    //Cyclic task index is invalid

#ifdef ECAT_DEBUG_EVENT_CALLBACKS
      LogError("ECAT-DEBUG: Cyclic task index is invalid");
#endif

//*******************************************************************************************************************************************************
    ECATM_EVTC_IOVAR_NO_DATA:
    //No input process image is available

#ifdef ECAT_DEBUG_EVENT_CALLBACKS
      LogError("ECAT-DEBUG: No input process image is available");
#endif

//*******************************************************************************************************************************************************
    ECATM_EVTC_IOVAR_BAD_CRC:
    //invalid crc

#ifdef ECAT_DEBUG_EVENT_CALLBACKS
      LogError("ECAT-DEBUG: invalid crc");
#endif

//*******************************************************************************************************************************************************
    ECATM_EVTC_MST_NO_ENICFG:
    //No ENI configuration loaded

#ifdef ECAT_DEBUG_EVENT_CALLBACKS
      LogError("ECAT-DEBUG: No ENI configuration loaded");
#endif

//*******************************************************************************************************************************************************
    ECATM_EVTC_MST_ENI_LOADED:
    //ENI shall get linked while another ENI configuration is still linked

#ifdef ECAT_DEBUG_EVENT_CALLBACKS
      LogError("ECAT-DEBUG: ENI shall get linked while another ENI configuration is still linked");
#endif

//*******************************************************************************************************************************************************
    ECATM_EVTC_MST_ACTIVATED:
    //Master is activated

#ifdef ECAT_DEBUG_EVENT_CALLBACKS
      LogError("ECAT-DEBUG: Master activated");
      LogValue("ECAT-DEBUG:Master activated after 0x{0}ms", (ops.tAbsolute-udInitStartTime));
#endif

//*******************************************************************************************************************************************************
    ECATM_EVTC_MST_DEACTIVATED:
    //Master is deactivated

#ifdef ECAT_DEBUG_EVENT_CALLBACKS
      LogError("ECAT-DEBUG: Master deactivated");
#endif

//*******************************************************************************************************************************************************
    ECATM_EVTC_MST_STATE_CHANGE:
    //Master ESM transition succeeded
    //arg1 ... old state
    //arg2 ... new state

#ifdef ECAT_DEBUG_EVENT_CALLBACKS
      LogValue("ECAT-DEBUG: Master State transition succeeded. Old State: 0x{0}, New State: 0x{1}", evt^.arg1$UDINT, evt^.arg2$UDINT);
#endif

      if evt^.arg2$t_e_ECAT_STATE <= ECAT_STATE_INIT then
        _SyncMeasureECAT1.Reset_Measurement();
      end_if;

      NewMasterEtherCATState := evt^.arg2$t_e_ECAT_STATE;

//*******************************************************************************************************************************************************
    ECATM_EVTC_MST_TRANS_FAILED:
    //Master ESM transition failed

#ifdef ECAT_DEBUG_EVENT_CALLBACKS
      LogValue("ECAT-DEBUG: Master State transition failed. State transition: 0x{0} to 0x{1}, error code: 0x{2}", evt^.arg1$UDINT, evt^.arg2$UDINT,evt^.arg3$UDINT);
#endif

      //Error during initialisation
      if bd_Flags.bPostInitFinished = FALSE then
        ErrorInitStep := InitSSW;
        InitSSW := _PrepareError;
        ClassState := _ManagerError;
        EtherCATState := ECAT_STATE_NONE;
      else
        if bd_Flags.bIsRequired then
          SetRequiredError( bLogInMethAllowed := bLogInCallbackAllowed);
        end_if;
      end_if;

//*******************************************************************************************************************************************************
    ECATM_EVTC_MST_ACTIVATE_ERR:
    //Master activation request failed. Master is de-activated.

#ifdef ECAT_DEBUG_EVENT_CALLBACKS
      LogError("ECAT-DEBUG: Master activation request failed. Master is de-activated.");
#endif

//*******************************************************************************************************************************************************

    ECATM_EVTC_MST_ESM_TMO:
    //Timeout for the synchronization of the acyclic task and the cyclic tasks during an ESM
    //transition. See also the transition flag ECATM_TRANS_IGNORE_WKC_SO.

#ifdef ECAT_DEBUG_EVENT_CALLBACKS
      LogError("ECAT-DEBUG: Timeout for the synchronization of the acyclic task and the cyclic tasks during an ESM transition");
#endif

//*******************************************************************************************************************************************************
    ECATM_EVTC_SLV_STATE_CHANGE:
    //Slave ESM transition succeeded

#ifdef ECAT_DEBUG_EVENT_CALLBACKS
      LogValue("ECAT-DEBUG: Slave State of Slave 0x{0} changed. Old State: 0x{1}, New State: 0x{2}", evt^.arg1$UDINT, evt^.arg2$UDINT, evt^.arg3$UDINT);
#endif

      //Forward callback to slave
      SendEvtCallBacktoSlave(udMasterID, evt, EventType, uiCallbackInfo);

//*******************************************************************************************************************************************************
    ECATM_EVTC_SLV_TRANS_FAILED:
    //Slave ESM transition failed

#ifdef ECAT_DEBUG_EVENT_CALLBACKS
      LogValue("ECAT-DEBUG: Slave State transition of Slave 0x{0} failed. Old State: 0x{1}, New State: 0x{2}", evt^.arg1$UDINT, evt^.arg2$UDINT, evt^.arg3$UDINT);
      LogValue("ECAT-DEBUG: Error Event Code: 0x{0} ", evt^.arg4$UDINT);
#endif

      //Forward callback to slave
      SendEvtCallBacktoSlave(udMasterID, evt, EventType, uiCallbackInfo);

      if evt^.arg1$UDINT <= sSlaveInfo.udMaxSlaves then
        pCurrentSlave := sSlaveInfo.pSlaves + (evt^.arg1$UDINT * sizeof(t_sSlaveInfo));

        //Check if slave was required
        if pCurrentSlave^.bRequired = TRUE then

          if bLogInCallbackAllowed then
            LogValue("@0575 (ECAT_Master_Base::EvtCallBack) State transition of required Slave 0x{0} failed.",evt^.arg1$UDINT);
          else
            bd_LogRtMessagesInCy.PostIt.SlvTransFailed := TRUE;
            bd_LogRtMessagesInCy.aLogValue1[5]         := evt^.arg1$UDINT;
          end_if;

          SetRequiredError( pTargetThis       := pCurrentSlave^.pThis
                          , udSlaveIndex      := pCurrentSlave^.udSlaveIndex
                          , bLogInMethAllowed := bLogInCallbackAllowed);

        elsif sDCInfo.DCModuleEnabled = TRUE & pCurrentSlave^.udSlaveIndex = sDCInfo.udSlaveIndex then

          if bLogInCallbackAllowed then
            LogValue("@0580 (ECAT_Master_Base::EvtCallBack) State transition of DC Module 0x{0} failed.",evt^.arg1$UDINT);
          else
            bd_LogRtMessagesInCy.PostIt.DCSlaveTransFailed := TRUE;
            bd_LogRtMessagesInCy.aLogValue1[15]         := evt^.arg1$UDINT;
          end_if;

          //DC Module is active but transition failed --> Set master into an error state
          ClassState := _ManagerError;
          EtherCATState := ECAT_STATE_NONE;
          InitSSW := _PrepareError;

        end_if;

          // Loggin else already done in SendEvtCallBacktoSlave
//      else
//        //Invalid slave no

      end_if;

//*******************************************************************************************************************************************************
    ECATM_EVTC_SLV_ACKERR_FAILED:
    //Slave error indication acknowledgment failed

#ifdef ECAT_DEBUG_EVENT_CALLBACKS
      LogValue("ECAT-DEBUG: Slave error indication acknowledgment failed. Slave Index 0x{0}, ErrorCode: 0x{1}", evt^.arg1$UDINT, evt^.arg2$UDINT);
#endif

      //Forward callback to slave
      SendEvtCallBacktoSlave(udMasterID, evt, EventType, uiCallbackInfo);

//*******************************************************************************************************************************************************
    ECATM_EVTC_ESM_BAD_CUR_STATE:
    //State request failed because of bad current state

#ifdef ECAT_DEBUG_EVENT_CALLBACKS
      LogError("ECAT-DEBUG: State request failed because of bad current state.");
#endif

//*******************************************************************************************************************************************************
    ECATM_EVTC_ESM_BAD_REQ_STATE:
    //Requested state does not exist

#ifdef ECAT_DEBUG_EVENT_CALLBACKS
      LogError("ECAT-DEBUG: Requested state does not exist.");
#endif

//*******************************************************************************************************************************************************
    ECATM_EVTC_ESM_REQ_BUSY:
    //ESM is currently performing a transition

#ifdef ECAT_DEBUG_EVENT_CALLBACKS
      LogError("ECAT-DEBUG: ESM is currently performing a transition.");
#endif
//*******************************************************************************************************************************************************
    ECATM_EVTC_INITC_RCV_TMO:
    //Init command failed with frame timeout error

    //arg1 ... device index: int
    //arg2 ... init cmd id: int

#ifdef ECAT_DEBUG_EVENT_CALLBACKS
      LogValue("ECAT-DEBUG: Init command failed with frame timeout error. Device Index: 0x{0}, Init cmd id: 0x{1}",evt^.arg1$UDINT, evt^.arg2$UDINT);
#endif

      //Forward callback to slave
      if evt^.arg1 >= 0 then  // device index -1 = Master
        SendEvtCallBacktoSlave(udMasterID, evt, EventType, uiCallbackInfo);
      end_if;

      if bLogInCallbackAllowed then
        LogValue("@057B (ECAT_Master_Base::EvtCallBack) Init command failed with frame timeout error. Device Index: 0x{0}, Init cmd id: 0x{1}",evt^.arg1$UDINT, evt^.arg2$UDINT);
      else
        bd_LogRtMessagesInCy.PostIt.InitCRecvTimeout  := TRUE;
        bd_LogRtMessagesInCy.aLogValue1[10]           := evt^.arg1$UDINT;
      end_if;

      if (evt^.arg1 >= 0) & (evt^.arg1$UDINT <= sSlaveInfo.udMaxSlaves) then
        pCurrentSlave := sSlaveInfo.pSlaves + (evt^.arg1$UDINT * sizeof(t_sSlaveInfo));

        //Check if slave was required
        if pCurrentSlave^.bRequired = TRUE then

          SetRequiredError( pTargetThis       := pCurrentSlave^.pThis
                          , udSlaveIndex      := pCurrentSlave^.udSlaveIndex
                          , bLogInMethAllowed := bLogInCallbackAllowed);
        end_if;

          // Loggin else already done in SendEvtCallBacktoSlave
//      else
//        //Invalid slave no

      end_if;

//*******************************************************************************************************************************************************
    ECATM_EVTC_INITC_VALID_WKC:
    //Init command failed with wrong working counter

    //arg1 ... device index: int
    //arg2 ... init cmd id: int
    //arg3 ... received WKC: int
    //arg4 ... expected WKC: int
    //txt ... Comment of init command in ENI file

#ifdef ECAT_DEBUG_EVENT_CALLBACKS
      LogValue("ECAT-DEBUG: Init command failed with wrong working counter. Device Index: 0x{0}",evt^.arg1$UDINT);
      LogValue("ECAT-DEBUG: init cmd id: 0x{0}, received WKC: 0x{1}, expected WKC: 0x{2}",evt^.arg2$UDINT, evt^.arg3$UDINT, evt^.arg4$UDINT);
      LogError(#evt^.txt[0]);
#endif

      if evt^.arg1 = -1 then  // If Master
        ClassState := _WrongHardware;
      end_if;

      //Forward callback to slave
      if evt^.arg1 >= 0 then // device index -1 = Master
        SendEvtCallBacktoSlave(udMasterID, evt, EventType, uiCallbackInfo);
      end_if;

      if bLogInCallbackAllowed then
        if evt^.arg1 = -1 then  // If Master
          LogError("@057C (ECAT_Master_Base::EvtCallBack) Init command failed with wrong working counter. Device: Master");
        else
          LogValue("@057C (ECAT_Master_Base::EvtCallBack) Init command failed with wrong working counter. Device Index: 0x{0}",evt^.arg1$UDINT);
        end_if;
        LogValue("@057C: init cmd id: 0x{0}, received WKC: 0x{1}, expected WKC: 0x{2}",evt^.arg2$UDINT, evt^.arg3$UDINT, evt^.arg4$UDINT);
        HWC_LogPrintf(pThis:=this, format:="@057C: %s", p0:=#evt^.txt[0]);
      else
        bd_LogRtMessagesInCy.PostIt.InitCValidWKC   := TRUE;
        bd_LogRtMessagesInCy.aLogValue1[11]         := evt^.arg1$UDINT;
      end_if;

      if (evt^.arg1 >= 0) & (evt^.arg1$UDINT <= sSlaveInfo.udMaxSlaves) then
        pCurrentSlave := sSlaveInfo.pSlaves + (evt^.arg1$UDINT * sizeof(t_sSlaveInfo));

        //Check if slave was required
        if pCurrentSlave^.bRequired = TRUE then

          SetRequiredError( pTargetThis       := pCurrentSlave^.pThis
                          , udSlaveIndex      := pCurrentSlave^.udSlaveIndex
                          , bLogInMethAllowed := bLogInCallbackAllowed);
        end_if;

          // Loggin else already done in SendEvtCallBacktoSlave
//      else
//        //Invalid slave no

      end_if;

//*******************************************************************************************************************************************************
    ECATM_EVTC_INITC_VALID_LEN:
    //Init command failed with invalid frame length

    //arg1 ... device index: int
    //arg2 ... init cmd id: int
    //arg3 ... received length
    //arg4 ... expected length
    //txt ... Comment of init command in ENI file

#ifdef ECAT_DEBUG_EVENT_CALLBACKS
      LogValue("ECAT-DEBUG: Init command failed with invalid frame length. Device Index: 0x{0}",evt^.arg1$UDINT);
      LogValue("ECAT-DEBUG: init cmd id: 0x{0}, received length: 0x{1}, expected length: 0x{2}",evt^.arg2$UDINT, evt^.arg3$UDINT, evt^.arg4$UDINT);
      LogError(#evt^.txt[0]);
#endif

      //Forward callback to slave
      if evt^.arg1 >= 0 then // device index -1 = Master
        SendEvtCallBacktoSlave(udMasterID, evt, EventType, uiCallbackInfo);
      end_if;

      if bLogInCallbackAllowed then
        LogValue("@09C8 (ECAT_Master_Base::EvtCallBack) Init command failed with invalid frame length. Device Index: 0x{0}",evt^.arg1$UDINT);
        LogValue("@09C8: init cmd id: 0x{0}, received length: 0x{1}, expected length: 0x{2}",evt^.arg2$UDINT, evt^.arg3$UDINT, evt^.arg4$UDINT);
        HWC_LogPrintf(pThis:=this, format:="@09C8: %s", p0:=#evt^.txt[0]);
      else
        bd_LogRtMessagesInCy.PostIt.InitCValidLen := TRUE;
        bd_LogRtMessagesInCy.aLogValue1[12]         := evt^.arg1$UDINT;
      end_if;

      if (evt^.arg1 >= 0) & (evt^.arg1$UDINT <= sSlaveInfo.udMaxSlaves) then
        pCurrentSlave := sSlaveInfo.pSlaves + (evt^.arg1$UDINT * sizeof(t_sSlaveInfo));

        //Check if slave was required
        if pCurrentSlave^.bRequired = TRUE then

          SetRequiredError( pTargetThis       := pCurrentSlave^.pThis
                          , udSlaveIndex      := pCurrentSlave^.udSlaveIndex
                          , bLogInMethAllowed := bLogInCallbackAllowed);
        end_if;

          // Loggin else already done in SendEvtCallBacktoSlave
//      else
//        //Invalid slave no

      end_if;

//*******************************************************************************************************************************************************
    ECATM_EVTC_INITC_VALID_DATA:
    //Init command failed during data validation

    //arg1 ... device index: int
    //arg2 ... init cmd id: int
    //arg3 ... byte index: int
    //arg4 ... received byte: uint8_t
    //txt ... Comment of init command in ENI file

#ifdef ECAT_DEBUG_EVENT_CALLBACKS
      LogValue("ECAT-DEBUG: Init command failed during data validation. Device Index: 0x{0}",evt^.arg1$UDINT);
      LogValue("ECAT-DEBUG: init cmd id: 0x{0}, byte index: 0x{1}, received byte: 0x{2}",evt^.arg2$UDINT, evt^.arg3$UDINT, evt^.arg4$UDINT);
      LogError(#evt^.txt[0]);
#endif

      //Forward callback to slave
      if evt^.arg1 >= 0 then  // device index -1 = Master
        SendEvtCallBacktoSlave(udMasterID, evt, EventType, uiCallbackInfo);
      end_if;

      if bLogInCallbackAllowed then
        LogValue("@057E (ECAT_Master_Base::EvtCallBack) Init command failed during data validation. Device Index: 0x{0}",evt^.arg1$UDINT);
        LogValue("@057E init cmd id: 0x{0}, byte index: 0x{1}, received byte: 0x{2}",evt^.arg2$UDINT, evt^.arg3$UDINT, evt^.arg4$UDINT);
        HWC_LogPrintf(pThis:=this, format:="@057E: %s", p0:=#evt^.txt[0]);
      else
        bd_LogRtMessagesInCy.PostIt.InitCValidData := TRUE;
        bd_LogRtMessagesInCy.aLogValue1[13]         := evt^.arg1$UDINT;
      end_if;

      if (evt^.arg1 >= 0) & (evt^.arg1$UDINT <= sSlaveInfo.udMaxSlaves) then
        pCurrentSlave := sSlaveInfo.pSlaves + (evt^.arg1$UDINT * sizeof(t_sSlaveInfo));

        //Check if slave was required
        if pCurrentSlave^.bRequired = TRUE then
          SetRequiredError( pTargetThis       := pCurrentSlave^.pThis
                          , udSlaveIndex      := pCurrentSlave^.udSlaveIndex
                          , bLogInMethAllowed := bLogInCallbackAllowed);
        end_if;

        // Loggin else already done in SendEvtCallBacktoSlave
//      else
//        //Invalid slave no

      end_if;

//*******************************************************************************************************************************************************
    ECATM_EVTC_MBX_BAD_RSP_MBXHD:
    //Bad mailbox header received

    //arg1 ... slave index: int

#ifdef ECAT_DEBUG_EVENT_CALLBACKS
      LogValue("ECAT-DEBUG: Bad mailbox header received. SlaveIndex: 0x{0}",evt^.arg1$UDINT);
#endif

//*******************************************************************************************************************************************************
    ECATM_EVTC_MBX_WR_FAILED:
    //Mailbox write failed due to invalid response

#ifdef ECAT_DEBUG_EVENT_CALLBACKS
      LogError("ECAT-DEBUG: Mailbox write failed due to invalid response.");
#endif

//*******************************************************************************************************************************************************
    ECATM_EVTC_MBX_RD_REPEAT_FAIL:
    //Mailbox read repeat counter reached

    //arg1 ... slave index: int

#ifdef ECAT_DEBUG_EVENT_CALLBACKS
      LogValue("ECAT-DEBUG: Mailbox read repeat counter reached. SlaveIndex: 0x{0}",evt^.arg1$UDINT);
#endif

//*******************************************************************************************************************************************************
    ECATM_EVTC_MBX_WR_REPEAT_FAIL:
    //Mailbox write repeat counter reached

#ifdef ECAT_DEBUG_EVENT_CALLBACKS
      LogError("ECAT-DEBUG: Mailbox write repeat counter reached.");
#endif

//*******************************************************************************************************************************************************
    ECATM_EVTC_MBX_RD_FAILED:
    //Mailbox read failed due to invalid response

    //arg1 ... slave index: int

#ifdef ECAT_DEBUG_EVENT_CALLBACKS
      LogValue("ECAT-DEBUG: Mailbox read failed due to invalid response. SlaveIndex: 0x{0}",evt^.arg1$UDINT);
#endif

//*******************************************************************************************************************************************************
    ECATM_EVTC_MBX_ERR_UNKNOWN_PROT:
    //Mailbox response with unknown protocol received

#ifdef ECAT_DEBUG_EVENT_CALLBACKS
      LogError("ECAT-DEBUG: Mailbox response with unknown protocol received.");
#endif

//*******************************************************************************************************************************************************
    ECATM_EVTC_MBX_ERR_REPLY:
    //Slave sent mailbox protocol error

    //arg1 ... slave index: int
    //arg2 ... type: int
    //arg3 ... detail: int

#ifdef ECAT_DEBUG_EVENT_CALLBACKS
      LogValue("ECAT-DEBUG: Slave sent mailbox protocol error. SlaveIndex: 0x{0}, type: 0x{1}, detail: 0x{2}",evt^.arg1$UDINT, evt^.arg2$UDINT, evt^.arg3$UDINT);
#endif

//*******************************************************************************************************************************************************
    ECATM_EVTC_COE_BAD_RSP:
    //Bad CoE response received

    //arg1 ... slave index: int

#ifdef ECAT_DEBUG_EVENT_CALLBACKS
      LogValue("ECAT-DEBUG: Bad CoE response received. SlaveIndex: 0x{0}",evt^.arg1$UDINT);
#endif

//*******************************************************************************************************************************************************
    ECATM_EVTC_COE_SDO_TRF_ERR:
    //CoE transfer error detected

    //arg1 ... slave index: int
    //arg2 ... index: uint16_t
    //arg3 ... subidx : uint8_t
    //arg4 ... error event code: int

    //  Ignore bLogInCallbackAllowed = FALSE, COE_SDO Event are always LSL_ECATM_ACYCLIC_TASK
    if bLogInCallbackAllowed & (EtherCATState < ECAT_STATE_OP) then // Log if < ECAT_STATE_OP, probably Init Cmd failed which are not handled in the Slave HW-Classes

      LogValue("@09B3 (ECAT_Master_Base::EvtCallBack) CoE transfer error detected. SlaveIndex: 0x{0}",evt^.arg1$UDINT);
      LogValue("@09B3 index: 0x{0}, subidx: 0x{1}, error event code: 0x{2}",evt^.arg2$UDINT, evt^.arg3$UDINT, evt^.arg4$UDINT);

#ifdef ECAT_DEBUG_EVENT_CALLBACKS
    else
      LogValue("ECAT-DEBUG: CoE transfer error detected. SlaveIndex: 0x{0}",evt^.arg1$UDINT);
      LogValue("ECAT-DEBUG: index: 0x{0}, subidx: 0x{1}, error event code: 0x{2}",evt^.arg2$UDINT, evt^.arg3$UDINT, evt^.arg4$UDINT);
#endif
    end_if;

//*******************************************************************************************************************************************************
    ECATM_EVTC_COE_SDO_TRF_TMO:
    //CoE timeout error detected

    //arg1 ... slave index: int
    //arg2 ... index: uint16_t
    //arg3 ... subidx : uint8_t

    //  Ignore bLogInCallbackAllowed = FALSE, COE_SDO Event are always LSL_ECATM_ACYCLIC_TASK
    if bLogInCallbackAllowed & (EtherCATState < ECAT_STATE_OP) then // Log if < ECAT_STATE_OP, probably Init Cmd failed which are not handled in the Slave HW-Classes

      LogValue("@09B4 (ECAT_Master_Base::EvtCallBack) CoE timeout error detected. SlaveIndex: 0x{0}",evt^.arg1$UDINT);
      LogValue("@09B4 index: 0x{0}, subidx: 0x{1}",evt^.arg2$UDINT, evt^.arg3$UDINT);

#ifdef ECAT_DEBUG_EVENT_CALLBACKS
    else
      LogValue("ECAT-DEBUG: CoE timeout error detected. SlaveIndex: 0x{0}",evt^.arg1$UDINT);
      LogValue("ECAT-DEBUG: index: 0x{0}, subidx: 0x{1}",evt^.arg2$UDINT, evt^.arg3$UDINT);
#endif
    end_if;

//*******************************************************************************************************************************************************
    ECATM_EVTC_COE_SDO_UPL_BUFSIZE:
    //CoE upload failed because of invalid receive buffer size

    //arg1 ... slave index: int
    //arg2 ... index: uint16_t
    //arg3 ... subidx : uint8_t
    //arg4 ... required size: int

    //  Ignore bLogInCallbackAllowed = FALSE, COE_SDO Event are always LSL_ECATM_ACYCLIC_TASK
    if bLogInCallbackAllowed & (EtherCATState < ECAT_STATE_OP) then // Log if < ECAT_STATE_OP, probably Init Cmd failed which are not handled in the Slave HW-Classes

      LogValue("@09B5 (ECAT_Master_Base::EvtCallBack) CoE upload failed because of invalid receive buffer size. SlaveIndex: 0x{0}",evt^.arg1$UDINT);
      LogValue("@09B5 index: 0x{0}, subidx: 0x{1}, required size: 0x{2}",evt^.arg2$UDINT, evt^.arg3$UDINT, evt^.arg4$UDINT);

#ifdef ECAT_DEBUG_EVENT_CALLBACKS
    else
      LogValue("ECAT-DEBUG: CoE upload failed because of invalid receive buffer size. SlaveIndex: 0x{0}",evt^.arg1$UDINT);
      LogValue("ECAT-DEBUG: index: 0x{0}, subidx: 0x{1}, required size: 0x{2}",evt^.arg2$UDINT, evt^.arg3$UDINT, evt^.arg4$UDINT);
#endif
    end_if;

//*******************************************************************************************************************************************************
    ECATM_EVTC_COE_SDO_ABORT_REQ:
    //CoE abort code received

    //arg1 ... slave index: int
    //arg2 ... index: uint16_t
    //arg3 ... subidx : uint8_t
    //arg4 ... abort code: uint32_t

    //  Ignore bLogInCallbackAllowed = FALSE, COE_SDO Event are always LSL_ECATM_ACYCLIC_TASK
    if bLogInCallbackAllowed & (EtherCATState < ECAT_STATE_OP) then // Log if < ECAT_STATE_OP, probably Init Cmd failed which are not handled in the Slave HW-Classes

      LogValue("@09B6 (ECAT_Master_Base::EvtCallBack): CoE abort code received. SlaveIndex: 0x{0}",evt^.arg1$UDINT);
      LogValue("@09B6 index: 0x{0}, subidx: 0x{1}, abort code: 0x{2}",evt^.arg2$UDINT, evt^.arg3$UDINT, evt^.arg4$UDINT);

#ifdef ECAT_DEBUG_EVENT_CALLBACKS
    else
      LogValue("ECAT-DEBUG: CoE abort code received. SlaveIndex: 0x{0}",evt^.arg1$UDINT);
      LogValue("ECAT-DEBUG: index: 0x{0}, subidx: 0x{1}, abort code: 0x{2}",evt^.arg2$UDINT, evt^.arg3$UDINT, evt^.arg4$UDINT);
#endif
    end_if;

//*******************************************************************************************************************************************************
    ECATM_EVTC_COE_EMERGENCY_MSG:
    //CoE emergency received

    //arg1 ... slave index: int
    //arg2 ... error code (16bit); register (16bit)
    //arg3 ... data1_4: 4x uint8_t
    //arg4 ... data 0: uint8_t

#ifdef ECAT_DEBUG_EVENT_CALLBACKS
      LogValue("ECAT-DEBUG: CoE emergency received. SlaveIndex: 0x{0}",evt^.arg1$UDINT);
      LogValue("ECAT-DEBUG: ErrorCode: 0x{0}, Data1_4: 0x{1}, Data0: 0x{2}",evt^.arg2$UDINT, evt^.arg3$UDINT, evt^.arg4$UDINT);
#endif

//*******************************************************************************************************************************************************
    ECATM_EVTC_EOE_INITC_BAD_RSP:

    //Bad response received for an EoE initalizaton command
    //arg1 ... slave index: int
    //arg2 ... initalizaton command index: int
    //arg3 ... response error code: int

#ifdef ECAT_DEBUG_EVENT_CALLBACKS
      LogValue("ECAT-DEBUG: Bad response received for an EoE initalizaton command SlaveIndex: 0x{0}",evt^.arg1$UDINT);
      LogValue("ECAT-DEBUG: Init Command: 0x{0},ErrorCode : 0x{1}",evt^.arg2$UDINT, evt^.arg3$UDINT);
#endif

//*******************************************************************************************************************************************************
    ECATM_EVTC_EOE_MBX_TRF_ERR:

    //EoE send request failed with mailbox error
    //arg1 ... slave index: int
    //arg2 ... mailbox error :int

#ifdef ECAT_DEBUG_EVENT_CALLBACKS
      LogValue("ECAT-DEBUG: EoE send request failed with mailbox error SlaveIndex: 0x{0} MBxErrorCode: 0x{1}", evt^.arg1$UDINT, evt^.arg2$UDINT);

#endif

//*******************************************************************************************************************************************************
    ECATM_EVTC_EOE_INITC_TMO:

    //EoE initalizaton command timed out
    //arg1 ... slave index: int
    //arg2 ... number of the init command

#ifdef ECAT_DEBUG_EVENT_CALLBACKS
      LogValue("ECAT-DEBUG: EoE initalizaton command timed out. SlaveIndex: 0x{0} INITCMD: 0x{1}", evt^.arg1$UDINT, evt^.arg2$UDINT);

#endif

//*******************************************************************************************************************************************************
    ECATM_EVTC_FOE_TRF_TMO:

#ifdef ECAT_DEBUG_EVENT_CALLBACKS
      LogError("ECAT-DEBUG: The event ECATM_EVTC_FOE_TRF_TMO occured");
#endif

//*******************************************************************************************************************************************************
    ECATM_EVTC_FOE_BAD_RSP:

#ifdef ECAT_DEBUG_EVENT_CALLBACKS
      LogError("ECAT-DEBUG: The event ECATM_EVTC_FOE_BAD_RSP occured");
#endif

//*******************************************************************************************************************************************************
    ECATM_EVTC_FOE_BAD_FRAMENO:

#ifdef ECAT_DEBUG_EVENT_CALLBACKS
      LogError("ECAT-DEBUG: The event ECATM_EVTC_FOE_BAD_FRAMENO occured");
#endif

//*******************************************************************************************************************************************************
    ECATM_EVTC_FOE_MBX_TOOSMALL:

#ifdef ECAT_DEBUG_EVENT_CALLBACKS
      LogError("ECAT-DEBUG: The event ECATM_EVTC_FOE_MBX_TOOSMALL occured");
#endif

//*******************************************************************************************************************************************************
    ECATM_EVTC_FOE_PARAM:

#ifdef ECAT_DEBUG_EVENT_CALLBACKS
      LogError("ECAT-DEBUG: The event ECATM_EVTC_FOE_PARAM occured");
#endif

//*******************************************************************************************************************************************************

//*******************************************************************************************************************************************************
    ECATM_EVTC_FRM_RCV_Q_EMPTY:
    //No free receive frame buffer (check ecatm configuration)

#ifdef ECAT_DEBUG_EVENT_CALLBACKS
      LogError("ECAT-DEBUG: No free receive frame buffer (check ecatm configuration)");
#endif

      ClassState := _InvalidConfguration;
      EtherCATState := ECAT_STATE_NONE;

      if bLogInCallbackAllowed then
        LogError("@0583 (ECAT_Master_Base::EvtCallBack) No free receive frame buffer (check ecatm configuration)");
      else
        bd_LogRtMessagesInCy.PostIt.NoFreeReceiveFrameBuffer := TRUE;
      end_if;

//*******************************************************************************************************************************************************
    ECATM_EVTC_FRM_RCV_LEN_TOO_BIG:
    //Too large EtherCAT frame received

    //arg1 ... frame size : int
    //arg2 ... descriptor size : int

#ifdef ECAT_DEBUG_EVENT_CALLBACKS
      LogValue("ECAT-DEBUG: Too large EtherCAT frame received. Framesize: 0x{0}, Descriptor Size: 0x{1}", evt^.arg1$UDINT, evt^.arg2$UDINT);
#endif

//*******************************************************************************************************************************************************
    ECATM_EVTC_FRM_RCV_BAD_LEN:
    //Received length doesn't match send length

    //arg1 ... received length: int
    //arg2 ... send length : int

#ifdef ECAT_DEBUG_EVENT_CALLBACKS
      LogValue("ECAT-DEBUG: Received length doesn't match send length . received length: 0x{0}, send length: 0x{1}", evt^.arg1$UDINT, evt^.arg2$UDINT);
#endif

//*******************************************************************************************************************************************************
    ECATM_EVTC_FRM_RCV_BAD_TYPE:
    //Received EtherCAT frame with bad type

    //arg1 ... type : uint8_t

#ifdef ECAT_DEBUG_EVENT_CALLBACKS
      LogValue("ECAT-DEBUG: Received EtherCAT frame with bad type . type: 0x{0}", evt^.arg1$UDINT);
#endif

//*******************************************************************************************************************************************************
    ECATM_EVTC_FRM_BAD_RSP_PDU:
    //Received PDU information does not match sent

    //arg1 ... byte index: int
    //arg2 ... send byte: uint8_t
    //arg3 ... received byte: uint8_t

#ifdef ECAT_DEBUG_EVENT_CALLBACKS
      LogValue("ECAT-DEBUG: Received length doesn't match send length . byte index: 0x{0}, send byte: 0x{1}, received: 0x{2}", evt^.arg1$UDINT, evt^.arg2$UDINT, evt^.arg3$UDINT);
#endif

//*******************************************************************************************************************************************************
    ECATM_EVTC_FRM_BAD_RSP_WKC:
    //Invalid Working counter received

#ifdef ECAT_DEBUG_EVENT_CALLBACKS
      LogError("ECAT-DEBUG: Invalid Working counter received");
#endif

//*******************************************************************************************************************************************************
    ECATM_EVTC_FRM_FULL:
    //Acyclic frame is full (PDUs must be sent in next loop)

#ifdef ECAT_DEBUG_EVENT_CALLBACKS
      LogError("ECAT-DEBUG: Acyclic frame is full (PDUs must be sent in next loop) ");
#endif

//*******************************************************************************************************************************************************
    ECATM_EVTC_FRM_BAD_CMD:
    //Invalid PDU command

#ifdef ECAT_DEBUG_EVENT_CALLBACKS
      LogError("ECAT-DEBUG: Invalid PDU command");
#endif

//*******************************************************************************************************************************************************
    ECATM_EVTC_FRM_NO_RCV:
    //Response frame timeout error

#ifdef ECAT_DEBUG_EVENT_CALLBACKS
      LogError("ECAT-DEBUG: Response frame timeout error");
#endif

//*******************************************************************************************************************************************************
    ECATM_EVTC_CFG_MAX_SIZE:
    //The configured maximum frame size _ecatm_cfg.frmsizemax is too small for a ESM initcmd,
    //a slave mailbox or a cyclic frame.
    //arg1 ... configured frame size (should be equal to _ecatm_cfg.frmsizemax): int
    //arg2 ... required frame size of the ENI: int

#ifdef ECAT_DEBUG_EVENT_CALLBACKS
      LogValue("ECAT-DEBUG: configured maximum frame size _ecatm_cfg.frmsizemax is too small. ConfSize: 0x{0}, reqiredSize: 0x{1}", evt^.arg1$UDINT, evt^.arg2$UDINT);
#endif

//*******************************************************************************************************************************************************
    ECATM_EVTC_LLETH_ERR:
    //Link layer error occurred (see ethll.h)

    //arg1 ... link layer error code: uint32_t

#ifdef ECAT_DEBUG_EVENT_CALLBACKS
      LogValue("ECAT-DEBUG: Link layer error occurred. Error code: 0x{0}", evt^.arg1$UDINT);
#endif

//*******************************************************************************************************************************************************
    ECATM_EVTC_LLETH_RCV_TMO:
    //Link layer frame receive timeout

#ifdef ECAT_DEBUG_EVENT_CALLBACKS
      LogError("ECAT-DEBUG: Link layer frame receive timeout");
#endif

//*******************************************************************************************************************************************************
    ECATM_EVTC_LLETH_FRM_NOTSENT:
    //Internal error code: Link layer failed to send a TX frame. The frame is still owned by the
    //hardware and shall not be altered.

#ifdef ECAT_DEBUG_EVENT_CALLBACKS
      LogError("ECAT-DEBUG: Event ECATM_EVTC_LLETH_FRM_NOTSENT occured");
#endif

//*******************************************************************************************************************************************************
    ECATM_EVTC_LLETH_LD_FRM_NOTSENT:
    //Internal error code: Link layer failed to send a TX frame and link is down. The frame is still
    //owned by the hardware and shall not be altered.

#ifdef ECAT_DEBUG_EVENT_CALLBACKS
      LogError("ECAT-DEBUG: Event ECATM_EVTC_LLETH_LD_FRM_NOTSENT occured");
#endif
//*******************************************************************************************************************************************************
    ECATM_EVTC_LLETH_LINK_DOWN:
    //Link layer link down detected

      DisconnectEvent(udMasterID:=udMasterID, evt:=evt, EventType:=EventType, uiCallbackInfo:=uiCallbackInfo);

#ifdef ECAT_DEBUG_EVENT_CALLBACKS
      LogError("ECAT-DEBUG: Link layer link down detected");
#endif

//*******************************************************************************************************************************************************
    ECATM_EVTC_LLETH_RX_REARM:
    //Re-arming frame at link layer failed

#ifdef ECAT_DEBUG_EVENT_CALLBACKS
      LogError("ECAT-DEBUG: Re-arming frame at link layer failed ");
#endif

//*******************************************************************************************************************************************************
    ECATM_EVTC_MON_ERR_TCP:
    //Monitor TCP stack error

#ifdef ECAT_DEBUG_EVENT_CALLBACKS
      LogError("ECAT-DEBUG: Monitor TCP stack error");
#endif

//*******************************************************************************************************************************************************
    ECATM_EVTC_MON_ERR_CONN:
    //Monitor TCP connection failed

#ifdef ECAT_DEBUG_EVENT_CALLBACKS
      LogError("ECAT-DEBUG: Monitor TCP connection failed ");
#endif

//*******************************************************************************************************************************************************
    ECATM_EVTC_MON_ERR_BAD_MSG:
    //Monitor: invalid message received

#ifdef ECAT_DEBUG_EVENT_CALLBACKS
      LogError("ECAT-DEBUG: invalid message received");
#endif

//*******************************************************************************************************************************************************
    ECATM_EVTC_MON_ERR_MSGBUFSIZE:
    //Monitor: invalid message buffer size

#ifdef ECAT_DEBUG_EVENT_CALLBACKS
      LogError("ECAT-DEBUG: invalid message buffer size ");
#endif

//*******************************************************************************************************************************************************
    ECATM_EVTC_MON_ERR_VERCHECK:
    //Monitor version does not match server version

#ifdef ECAT_DEBUG_EVENT_CALLBACKS
      LogError("ECAT-DEBUG: Monitor version does not match server version");
#endif

//*******************************************************************************************************************************************************
    ECATM_EVTC_SUP_SLV_NUM_CHG:
    //Supervision detected that slave number in network changed

#ifdef ECAT_DEBUG_EVENT_CALLBACKS
      LogError("ECAT-DEBUG: Supervision detected that slave number in network changed");
#endif

//*******************************************************************************************************************************************************
    ECATM_EVTC_SUP_SLV_STATE_CHG:
    //Supervision detected unexpected slave state change or error indication flag

#ifdef ECAT_DEBUG_EVENT_CALLBACKS
      LogError("ECAT-DEBUG: Supervision detected unexpected slave state change or error indication flag");
#endif

    //Forward callback to slave
    SendEvtCallBacktoSlave(udMasterID, evt, EventType, uiCallbackInfo);

//*******************************************************************************************************************************************************
    ECATM_EVTC_SUP_SLV_ALSTATUS_CHG:
    //Supervision detected changed of AL-Status Code of a slave

#ifdef ECAT_DEBUG_EVENT_CALLBACKS
      LogValue("ECAT-DEBUG: Supervision detected changed of AL-Status Code of a slave. Slave Index 0x{0}, Current State: 0x{1}, AL-Status Code: 0x{2}", evt^.arg1$UDINT, evt^.arg2$UDINT,evt^.arg3$UDINT);
#endif

      //Forward callback to slave
      SendEvtCallBacktoSlave(udMasterID, evt, EventType, uiCallbackInfo);

//*******************************************************************************************************************************************************
    ECATM_EVTC_SUP_SLV_WKC_UNEXPECT:
    //More than one slave with same physical address detected

#ifdef ECAT_DEBUG_EVENT_CALLBACKS
      LogError("ECAT-DEBUG: More than one slave with same physical address detected.");
#endif

//*******************************************************************************************************************************************************
    ECATM_EVTC_SUP_NET_REINIT_REQ:
    //Supervision failed to repair network. Re-initialization of network shall be done.

#ifdef ECAT_DEBUG_EVENT_CALLBACKS
      LogError("ECAT-DEBUG: Supervision failed to repair network. Re-initialization of network shall be done.");
#endif

//*******************************************************************************************************************************************************
    ECATM_EVTC_SUP_SLV_COMM_CHG:
    //Supervision detected that the slave connection status changed

#ifdef ECAT_DEBUG_EVENT_CALLBACKS
      LogValue("ECAT-DEBUG: Supervision detected that the slave connection status changed. Slvidx: 0x{0}, connected: 0x{1}, current state: 0x{2}", evt^.arg1$UDINT, evt^.arg2$UDINT, evt^.arg3$UDINT);
#endif

      //Forward callback to slave
      SendEvtCallBacktoSlave(udMasterID, evt, EventType, uiCallbackInfo);

//*******************************************************************************************************************************************************
    ECATM_EVTC_DC_MAX_RETRY:
    //DC step failed after max retries (frame loss or WKC error). The maximum number of retries is defined by CONFIG_ECATM_DC_MAXRETRY.
    //arg1 ... device index: slave index or ECATM_MST_DEVIDX

#ifdef ECAT_DEBUG_EVENT_CALLBACKS
      LogValue("ECAT-DEBUG: Event ECATM_EVTC_DC_MAX_RETRY occured. SlaveIndex = 0x{0}", evt^.arg1$UDINT);
#endif

//*******************************************************************************************************************************************************
    ECATM_EVTC_DC_SKIPPED:
    //Some configurators (e.g. TwinCAT 2) are marking each slave as DC slave.
    //The initialization of the slave failed and the master stack assumes that this slave doesn't require DC.
    //If this slave requires DC generate an error and request an INIT transition of the master.
    //arg1 ... slave index

#ifdef ECAT_DEBUG_EVENT_CALLBACKS
      LogValue("ECAT-DEBUG: Event ECATM_EVTC_DC_SKIPPED occured. SlaveIndex = 0x{0}", evt^.arg1$UDINT);
#endif

//*******************************************************************************************************************************************************
    ECATM_EVTC_DC_STATIC_DRIFT:
    //Static drift compensation failed with a timeout for the slave. ESM transition will fail with the error ECATM_EVTC_ESM_DC_FAILED.

#ifdef ECAT_DEBUG_EVENT_CALLBACKS
      LogValue("ECAT-DEBUG: Event ECATM_EVTC_DC_STATIC_DRIFT occured. SlaveIndex = 0x{0}", evt^.arg1$UDINT);
#endif

//*******************************************************************************************************************************************************
    ECATM_EVTC_DC_NOT_SUPPORTED:
    //A mandatory slave doesn't support DC (e.g. the reference slave or a multiple port slave)
    //arg1 ... slave index

#ifdef ECAT_DEBUG_EVENT_CALLBACKS
      LogValue("ECAT-DEBUG: Event ECATM_EVTC_DC_NOT_SUPPORTED occured. SlaveIndex = 0x{0}", evt^.arg1$UDINT);
#endif

//*******************************************************************************************************************************************************
    ECATM_EVTC_DC_REFSLAVE_32BIT:
    //The reference slave owns a 32-Bit counter for DC. The network time recovery is disabled. Change the network topology to fix this warning.
    //arg ... reference slave

#ifdef ECAT_DEBUG_EVENT_CALLBACKS
      LogValue("ECAT-DEBUG: Event ECATM_EVTC_DC_REFSLAVE_32BIT occured. SlaveIndex = 0x{0}", evt^.arg1$UDINT);
#endif

//*******************************************************************************************************************************************************
    ECATM_EVTC_DC_SET_SYNC:
    //The activation of the sync signal for this slave failed. Try to increase the _ecatm_dc_cfg.syncguardcycles to fix this error.
    //arg1 ... slave index

#ifdef ECAT_DEBUG_EVENT_CALLBACKS
      LogValue("ECAT-DEBUG: Event ECATM_EVTC_DC_SET_SYNC occured. SlaveIndex = 0x{0}", evt^.arg1$UDINT);
#endif

//*******************************************************************************************************************************************************
    ECATM_EVTC_DC_SYNC_WINDOW:
    //Slave was outside of the valid sync window during the last sync window refresh run. This event is only generated for the first time.
    //arg 1 ... slave index
    //arg 2 ... sync window: measured sync window of the slave

#ifdef ECAT_DEBUG_EVENT_CALLBACKS
      LogValue("ECAT-DEBUG: Event ECATM_EVTC_DC_SYNC_WINDOW occured. SlaveIndex = 0x{0}", evt^.arg1$UDINT);
#endif

//*******************************************************************************************************************************************************
    ECATM_EVTC_DC_FOUND:
    //Reference slave found during ecatm_eni_link(). DC module will be enabled.
    //arg1 ... slave index

#ifdef ECAT_DEBUG_EVENT_CALLBACKS
      LogValue("ECAT-DEBUG: Event ECATM_EVTC_DC_FOUND occured. SlaveIndex = 0x{0}", evt^.arg1$UDINT);
#endif

      sDCInfo.DCModuleEnabled  := TRUE;
      sDCInfo.udSlaveIndex     := evt^.arg1$UDINT;

      bs_Syncmodes.DC_Found := TRUE;

//*******************************************************************************************************************************************************
    ECATM_EVTC_DC_SYNC_DONE:
    //Static drift compensation finished. Slave will continue the its ESM transition.
    //arg1 ... slave index

    bs_Syncmodes.DC_Compensated := TRUE;

    _SyncMeasureECAT1.UpdateDCStatus(bs_Syncmodes);

#ifdef ECAT_DEBUG_EVENT_CALLBACKS
      LogValue("ECAT-DEBUG: Event ECATM_EVTC_DC_SYNC_DONE occured. SlaveIndex = 0x{0}", evt^.arg1$UDINT);
#endif

//*******************************************************************************************************************************************************
    ECATM_EVTC_DC_CYCLE_PERIOD:
    //The sync0 period of the slave is not a multiple or a fraction of the cyclic task period. The cyclic
    //task period is probably configured wrong or the slave is assigned to a sync unit of another
    //cyclic task (not supported by the master stack).
    //arg1 ... slave index

#ifdef ECAT_DEBUG_EVENT_CALLBACKS
      LogValue("ECAT-DEBUG: Event ECATM_EVTC_DC_CYCLE_PERIOD occured. SlaveIndex = 0x{0}", evt^.arg1$UDINT);
#endif

      ClassState := _InvalidConfguration;
      EtherCATState := ECAT_STATE_NONE;

      if bLogInCallbackAllowed then
        LogValue("@0581 (ECAT_Master_Base::EvtCallBack) Sync0 period of the slave 0x{0} is not a multiple or fraction of the cyclic task period",evt^.arg1$UDINT);
      else
        bd_LogRtMessagesInCy.PostIt.InvalidDCCyclePeriod := TRUE;
        bd_LogRtMessagesInCy.aLogValue1[16]              := evt^.arg1$UDINT;
      end_if;

//*******************************************************************************************************************************************************
    ECATM_EVTC_DC_SLV_OFFSET_REQ:
      //This event is generated during the IP transition of the master. The transition is held until the
    //function ecatm_dc_set_offset() is called.
    //Only Called in DC Slavemode
    //ECATM_EVTT_INFO
    //arg1   Link layer frame send timestamp: uint32_t
    //arg2   Link layer frame receive timestamp: uint32_t
    //arg3   Measured round trip time at the DC reference slave. The value is equal to the return
    //       value of _ecatm_dc_get_rtt(): uint32_t

    _syncmeasureECAT1.SetDCSlaveOffset(LLSend:= evt^.arg1$UDINT
                                   , LLReceive:= evt^.arg2$UDINT
                                      , DC_RTT:= evt^.arg3$UDINT);

#ifdef ECAT_DEBUG_EVENT_CALLBACKS
      LogError("ECAT-DEBUG: Event ECATM_EVTC_DC_SLV_OFFSET_REQ occured");
#endif

//*******************************************************************************************************************************************************
    ECATM_EVTC_DC_DISABLED:
      //DC disabled but refslave=%d found (DC slaves:%d)")
